(* IEC 61131-3 sources: Test-Git_ESME26/TestProgettoESME_26.fbsproj/PacDriveLib Migration/Motion/Homing/PDL_FB_HomeTp.fb.st^, 6 files *)

(* ---- EnableParameterCheck.meth.st ---- *)
METHOD PRIVATE EnableParameterCheck : BOOL
VAR
	xSuccess	: BOOL;
	ifGetParentDevice      : DTSI.IF_GetParentDevice;
	ifDeviceAccess         : DTSI.IF_DeviceAccess;
END_VAR

EnableParameterCheck := FALSE;
// querry all interfaces during enabeling
xSuccess := __QUERYINTERFACE(i_ifDrive, ifGetParentDevice);
IF NOT xSuccess OR ifGetParentDevice = 0 THEN
	SetDiagOutput(	i_etDiag	:= GD.ET_Diag.InputParameterInvalid,
					i_etDiagExt := PDL_ET_DiagExt.DriveInvalid,
					i_sMsg		:= 'i_ifDrive - IF_GetParentDevice not implemented.');
	RETURN;
END_IF
ifDeviceAccess := ifGetParentDevice.GetParentDevice();

xSuccess := __QUERYINTERFACE(ifDeviceAccess,ifScalingAccess );
IF (NOT xSuccess OR ifScalingAccess = 0) THEN
	SetDiagOutput(	i_etDiag	:= GD.ET_Diag.InputParameterInvalid,
					i_etDiagExt := PDL_ET_DiagExt.DriveInvalid,
					i_sMsg		:= 'i_ifDrive - IF_Scaling not implemented.');
	diState := 0;
	RETURN;
END_IF
ifScaling := ifScalingAccess.Scaling;

xSuccess := __QUERYINTERFACE(ifDeviceAccess,ifDrive2Access );
IF (NOT xSuccess OR ifDrive2Access = 0) THEN
	q_etDiag	:= GD.ET_Diag.InputParameterInvalid;
	q_etDiagExt := PDL_ET_DiagExt.DriveInvalid;
	q_sMsg		:= 'i_ifDrive - IF_Drive2 not implemented.';
	RETURN;
END_IF
ifDrive2 := ifDrive2Access.Drive2;

xSuccess := __QUERYINTERFACE(ifDeviceAccess,ifDriveAccess );
IF (NOT xSuccess OR ifDriveAccess = 0) THEN
	q_etDiag	:= GD.ET_Diag.InputParameterInvalid;
	q_etDiagExt := PDL_ET_DiagExt.DriveInvalid;
	q_sMsg		:= 'i_ifDrive - IF_Drive not implemented.';
	RETURN;
END_IF
ifDrive := ifDriveAccess.Drive;

xSuccess := __QUERYINTERFACE(ifDeviceAccess,ifDriveConfigAccess );
IF (NOT xSuccess OR ifDriveConfigAccess = 0) THEN
	SetDiagOutput(	i_etDiag	:= GD.ET_Diag.InputParameterInvalid,
					i_etDiagExt := PDL_ET_DiagExt.DriveInvalid,
					i_sMsg		:= 'i_ifDrive - IF_DriveConfig not implemented.');
	diState := 0;
	RETURN;
END_IF
ifDriveConfig := ifDriveConfigAccess.DriveConfig;

xSuccess := __QUERYINTERFACE(i_ifTouchProbe, ifGetParentDevice);
IF NOT xSuccess OR ifGetParentDevice = 0 THEN
	SetDiagOutput(	i_etDiag	:= GD.ET_Diag.InputParameterInvalid,
					i_etDiagExt := PDL_ET_DiagExt.DriveInvalid,
					i_sMsg		:= 'i_ifTouchProbe - IF_GetParentDevice not implemented.');
	RETURN;
END_IF
ifDeviceAccess := ifGetParentDevice.GetParentDevice();

xSuccess := __QUERYINTERFACE(ifDeviceAccess, ifTouprobeDataAccess);
IF NOT xSuccess OR (ifTouprobeDataAccess = 0) THEN
	SetDiagOutput(	i_etDiag	:= GD.ET_Diag.InputParameterInvalid,
					i_etDiagExt := PDL_ET_DiagExt.TouchProbeInvalid,
					i_sMsg		:= 'i_ifTouchProbe - IF_TouprobeDataAccess not implemented');
	RETURN;
END_IF
ifTouprobeData := ifTouprobeDataAccess.TouchprobeData;

xSuccess := __QUERYINTERFACE(ifDeviceAccess, ifDeviceTreeObjectAccess);
IF xSuccess THEN
	sDriveName := ifDeviceTreeObjectAccess.DeviceTreeObject.Name;
ELSE
	sDriveName := '';
END_IF

IF NOT StartParameterCheck() THEN
	; // parametrization fault -> diag message already set in StartParameterCheck()
ELSE
	fbSetPos.Axis           	:= i_ifDrive;

	fbStop.Axis 				:= i_ifDrive;
	fbStop.Deceleration 		:= i_lrDec;
	fbStop.Jerk 				:= i_lrJerk;

	fbMoveAbsolute.Axis    		:= i_ifDrive;
	fbMoveAbsolute.Velocity 	:= i_lrVel;
	fbMoveAbsolute.Deceleration := i_lrDec;
	fbMoveAbsolute.Acceleration := i_lrAcc;
	fbMoveAbsolute.Jerk 		:= i_lrJerk;
	fbMoveAbsolute.BufferMode	:= PLCO.MC_Buffer_Mode.Aborting;
	fbMoveAbsolute.Direction	:= PLCO.MC_Direction.PositiveDirection;

	fbMoveRelative.Axis     	:= i_ifDrive;
	fbMoveRelative.Velocity 	:= i_lrVel;
	fbMoveRelative.Deceleration := i_lrDec;
	fbMoveRelative.Acceleration := i_lrAcc;
	fbMoveRelative.Jerk 		:= i_lrJerk;
	fbMoveRelative.BufferMode	:= PLCO.MC_Buffer_Mode.Aborting;

	fbAbortTouchprobe.Axis  	:= i_ifDrive;
	fbAbortTouchprobe.ifTrigger	:= i_ifTouchProbe;

	fbTouchProbe.Axis 			:= i_ifDrive;
	fbTouchProbe.ifTrigger		:= i_ifTouchProbe;

	EnableParameterCheck := TRUE;
END_IF

(* ---- RegisterLoggerPoint.meth.st ---- *)
METHOD PUBLIC RegisterLoggerPoint
VAR_INPUT
	i_ifParent		: APL.IF_LoggerPoint;
	i_sName			: STRING[80];
END_VAR
VAR_OUTPUT
	q_etDiag		: GD.ET_Diag := GD.ET_Diag.Ok;
	q_etDiagExt		: PDL_ET_DiagExt := PDL_ET_DiagExt.Ok;
END_VAR
VAR
	etDiagBuffer		: GD.ET_Diag;
	etDiagExtBufferAPL	: APL.ET_DiagExt;
END_VAR

THIS^.fbLoggerPoint.RegisterLoggerPoint(	i_ifParent		:= i_ifParent,
											i_sName			:= i_sName,
											i_sType			:= 'FB_HomeTp',
											i_sSource		:= 'PDL',
											q_etDiag		=> etDiagBuffer,
											q_etDiagExt		=> etDiagExtBufferAPL);
IF (etDiagBuffer <> GD.ET_Diag.Ok) THEN
	CASE etDiagExtBufferAPL OF
		APL.ET_DiagExt.ParentInvalid:
			q_etDiag := GD.ET_Diag.InputParameterInvalid;
			q_etDiagExt := PDL_ET_DiagExt.ParentInvalid;

		APL.ET_DiagExt.ParentNotRegistered:
			q_etDiag := GD.ET_Diag.InputParameterInvalid;
			q_etDiagExt := PDL_ET_DiagExt.ParentNotRegistered;

		APL.ET_DiagExt.MaxNumberOfLoggerPointsExeeded:
			q_etDiag := GD.ET_Diag.InputParameterInvalid;
			q_etDiagExt := PDL_ET_DiagExt.MaxNumberOfLoggerPointsExeeded;

	ELSE
		q_etDiag := GD.ET_Diag.UnexpectedProgramBehavior;
		q_etdiagExt := PDL_ET_DiagExt.UnexpectedDiagExt;
	END_CASE
END_IF

(* ---- SetDiagOutput.meth.st ---- *)
METHOD PRIVATE SetDiagOutput
VAR_INPUT
	i_etDiag	: GD.ET_Diag;
	i_etDiagExt	: PDL_ET_DiagExt;
	i_sMsg		: STRING[80];
END_VAR
VAR
END_VAR

// check whether the new state can overwrite the current state
IF q_etDiag = GD.ET_Diag.OK OR i_etDiagExt = PDL_ET_DiagExt.Disabled THEN
	// set outputs
	q_etDiag 	:= i_etDiag;
	q_etDiagExt := i_etDiagExt;
	q_sMsg 		:= i_sMsg;
	IF (i_etDiag <> GD.ET_Diag.Ok) THEN
		q_xReady := FALSE;
	END_IF

	// set application logger entry
	IF(i_etDiag = GD.ET_Diag.Ok) AND (THIS^.fbLoggerPoint.etLogLevel >= APL.ET_LogLevel.StatusMessage) THEN
		THIS^.fbLoggerPoint.AddLogEntry(	i_etLogLevel	:= APL.ET_LogLevel.StatusMessage,
											i_etDiag		:= q_etDiag,
											i_udiDiagExt	:= q_etDiagExt,
											i_sMessage		:= SE_CTBX.FC_MultiConcat(	i_sString1	:= Standard.CONCAT('ET_Diag: ', GD.FC_EtDiagToString(q_etDiag)),
																						i_sString2	:= Standard.CONCAT(' PDL_ET_DiagExt: ', PDL_FC_EtDiagExtToString(q_etDiagExt)),
																						i_sString3	:= Standard.CONCAT(' sMsg: ', q_sMsg),
																						i_sString4	:= ''),
											q_etDiag		:= ,	// ignore result
											q_etDiagExt		:= );	// ignore result
	ELSIF(i_etDiag = GD.ET_Diag.UnexpectedProgramBehavior) AND (THIS^.fbLoggerPoint.etLogLevel >= APL.ET_LogLevel.CriticalException) THEN
		THIS^.fbLoggerPoint.AddLogEntry(	i_etLogLevel	:= APL.ET_LogLevel.CriticalException,
											i_etDiag		:= q_etDiag,
											i_udiDiagExt	:= q_etDiagExt,
											i_sMessage		:= SE_CTBX.FC_MultiConcat(	i_sString1	:= Standard.CONCAT('ET_Diag: ', GD.FC_EtDiagToString(q_etDiag)),
																						i_sString2	:= Standard.CONCAT(' PDL_ET_DiagExt: ', PDL_FC_EtDiagExtToString(q_etDiagExt)),
																						i_sString3	:= Standard.CONCAT(' sMsg: ', q_sMsg),
																						i_sString4	:= ''),
											q_etDiag		:= ,	// ignore result
											q_etDiagExt		:= );	// ignore result
	ELSE
		THIS^.fbLoggerPoint.AddLogEntry(	i_etLogLevel	:= APL.ET_LogLevel.Exception,
											i_etDiag		:= q_etDiag,
											i_udiDiagExt	:= q_etDiagExt,
											i_sMessage		:= SE_CTBX.FC_MultiConcat(	i_sString1	:= Standard.CONCAT('ET_Diag: ', GD.FC_EtDiagToString(q_etDiag)),
																						i_sString2	:= Standard.CONCAT(' PDL_ET_DiagExt: ', PDL_FC_EtDiagExtToString(q_etDiagExt)),
																						i_sString3	:= Standard.CONCAT(' sMsg: ', q_sMsg),
																						i_sString4	:= ''),
											q_etDiag		:= ,	// ignore result
											q_etDiagExt		:= );	// ignore result
	END_IF
END_IF

(* ---- SetTpEdge.meth.st ---- *)
METHOD PRIVATE SetTpEdge
VAR_INPUT
	i_xOppositeFlank	: BOOL;
END_VAR

IF i_etMode = PDL_ET_HomeTpMode.PosDirectionNegEdgeTp OR i_etMode = PDL_ET_HomeTpMode.NegDirectionNegEdgeTp THEN
	IF NOT i_xOppositeFlank THEN
		ifTouprobeData.CaptureEdgeSet := 0; // trigger on falling edge
	ELSE
		ifTouprobeData.CaptureEdgeSet := 1; // trigger on rising edge
	END_IF
ELSE
	IF NOT i_xOppositeFlank THEN
		ifTouprobeData.CaptureEdgeSet := 1; // trigger on rising edge
	ELSE
		ifTouprobeData.CaptureEdgeSet := 0; // trigger on falling edge
	END_IF
END_IF

(* ---- StartParameterCheck.meth.st ---- *)
METHOD PRIVATE StartParameterCheck : BOOL
VAR_INPUT
END_VAR

StartParameterCheck := FALSE;

IF i_ifDrive = 0 THEN
	SetDiagOutput(	i_etDiag	:= GD.ET_Diag.InputParameterInvalid,
					i_etDiagExt := PDL_ET_DiagExt.DriveInvalid,
					i_sMsg		:= 'i_ifDrive - Invalid Interface');
ELSIF i_ifTouchProbe = 0 THEN
	SetDiagOutput(	i_etDiag	:= GD.ET_Diag.InputParameterInvalid,
					i_etDiagExt := PDL_ET_DiagExt.TouchProbeInvalid,
					i_sMsg		:= 'i_ifTouchProbe - Invalid Interface');
ELSIF (i_lrMaxTravel <= 0.0) THEN
	SetDiagOutput(	i_etDiag	:= GD.ET_Diag.InputParameterInvalid,
					i_etDiagExt := PDL_ET_DiagExt.MaxTravelRange,
					i_sMsg		:= 'i_lrMaxTravel <= 0.0');
ELSIF i_lrVel <= 0.0  OR (ABS(i_lrVel) > ifDriveConfig.MaxVel AND ifDriveConfig.MaxVel <> 0) THEN
	SetDiagOutput(	i_etDiag	:= GD.ET_Diag.InputParameterInvalid,
					i_etDiagExt := PDL_ET_DiagExt.VelRange,
					i_sMsg		:= STANDARD.CONCAT('0.0 < i_lrVel <= ', TO_STRING(ifDriveConfig.MaxVel)) );
ELSIF i_lrAcc <= 0.0 OR (i_lrAcc > ifDriveConfig.MaxAcc AND ifDriveConfig.MaxAcc <> 0) THEN
	SetDiagOutput(	i_etDiag	:= GD.ET_Diag.InputParameterInvalid,
					i_etDiagExt := PDL_ET_DiagExt.AccRange,
					i_sMsg		:= STANDARD.CONCAT('0.0 < i_lrAcc <= ', TO_STRING(ifDriveConfig.MaxAcc) ));
ELSIF i_lrDec <= 0.0 OR (i_lrDec > ifDriveConfig.MaxAcc AND ifDriveConfig.MaxAcc <> 0)THEN
	SetDiagOutput(	i_etDiag	:= GD.ET_Diag.InputParameterInvalid,
					i_etDiagExt := PDL_ET_DiagExt.DecRange,
					i_sMsg		:= STANDARD.CONCAT('0.0 < i_lrDec <= ', TO_STRING(ifDriveConfig.MaxAcc) ));
ELSIF (i_etMode <> PDL_ET_HomeTpMode.PosDirectionPosEdgeTp) AND
	(i_etMode <> PDL_ET_HomeTpMode.NegDirectionPosEdgeTp) AND
	(i_etMode <> PDL_ET_HomeTpMode.NegDirectionNegEdgeTp) AND
	(i_etMode <> PDL_ET_HomeTpMode.PosDirectionNegEdgeTp) THEN
		SetDiagOutput(	i_etDiag	:= GD.ET_Diag.InputParameterInvalid,
						i_etDiagExt := PDL_ET_DiagExt.UnknownMode,
						i_sMsg		:= '');
ELSE
	lrDistance	:= i_lrMaxTravel;

	fbStop.Deceleration 		:= i_lrDec;
	fbStop.Jerk 				:= i_lrJerk;

	fbMoveAbsolute.Velocity 	:= i_lrVel;
	fbMoveAbsolute.Deceleration := i_lrDec;
	fbMoveAbsolute.Acceleration := i_lrAcc;
	fbMoveAbsolute.Jerk 		:= i_lrJerk;

	fbMoveRelative.Velocity 	:= i_lrVel;
	fbMoveRelative.Deceleration := i_lrDec;
	fbMoveRelative.Acceleration := i_lrAcc;
	fbMoveRelative.Jerk 		:= i_lrJerk;

	StartParameterCheck := TRUE;
END_IF

(* ---- StartPositioningAndTPEdge.meth.st ---- *)
METHOD PRIVATE StartPositioningAndTPEdge : BOOL
VAR_INPUT
	i_xOppositeDirection	: BOOL;
END_VAR
VAR
	lrDistance_loc		: LREAL;
END_VAR

IF
	(NOT i_xOppositeDirection AND (i_etMode = PDL_ET_HomeTpMode.PosDirectionNegEdgeTp OR i_etMode = PDL_ET_HomeTpMode.PosDirectionPosEdgeTp)) OR
	(i_xOppositeDirection AND (i_etMode = PDL_ET_HomeTpMode.NegDirectionNegEdgeTp OR i_etMode = PDL_ET_HomeTpMode.NegDirectionPosEdgeTp))
THEN
	lrDistance_loc := lrDistance;
ELSE
	lrDistance_loc := -lrDistance;
END_IF

xMotionJobStarted := FALSE;
fbMoveRelative(Execute := TRUE, Distance := lrDistance_loc);

IF fbMoveRelative.Error THEN
	SetDiagOutput(
		i_etDiag    := GD.ET_Diag.UnexpectedProgramBehavior,
		i_etDiagExt := PDL_ET_DiagExt.UnexpectedFeedback,
		i_sMsg      := CONCAT('MC_MoveRelative.ErrorID: ', PLCO.FC_EtResultToString(THIS^.fbMoveRelative.ErrorID))
	);
	THIS^.fbMoveRelative(Execute := FALSE);

ELSE
	q_xMotionInstructionActive := TRUE;
	fbTouchProbe(
		Execute       := TRUE,
		WindowOnly    := TRUE,
		FirstPosition := q_lrPosition - ABS(i_lrMaxTravel),
		LastPosition  := q_lrPosition + ABS(i_lrMaxTravel),
		PositionType  := PLCO.MC_PositionType.ActualPosition
	);

	IF fbTouchProbe.Error THEN
		SetDiagOutput(
			i_etDiag    := GD.ET_Diag.UnexpectedProgramBehavior,
			i_etDiagExt := PDL_ET_DiagExt.UnexpectedFeedback,
			i_sMsg      := CONCAT('MC_TouchProbe: ', PLCO.FC_EtResultToString(fbTouchProbe.ErrorId))
		);
		fbTouchProbe(Execute := FALSE);
	END_IF
	StartPositioningAndTPEdge := TRUE;
END_IF
